Fanuc TP program (LS listing): PgProg.LS

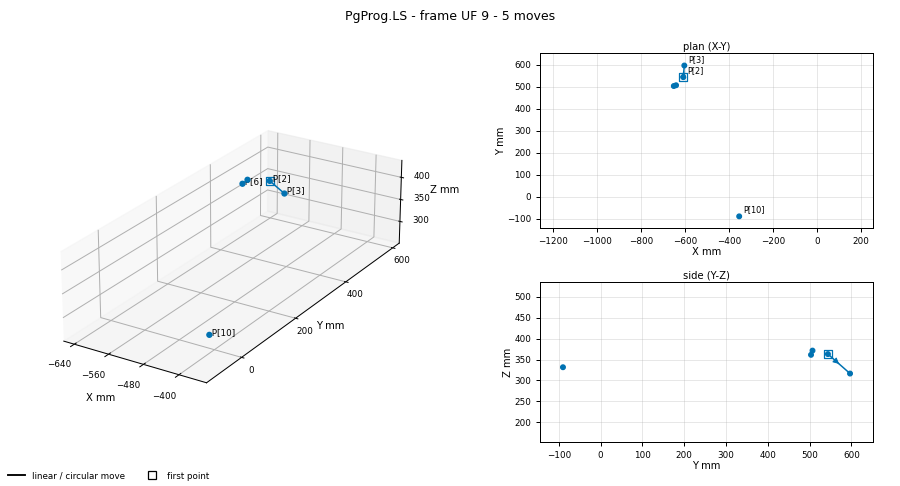
[picture p0: tool path of PgProg.LS in frame UF 9, 5 of 9 moves have a stored position in this frame; points joined in program order, loops and branches not executed]
/PROG  PgProg
/ATTR
OWNER		= MNEDITOR;
COMMENT		= "RoboDK sequence";
PROG_SIZE	= 0;
CREATE		= DATE 31-12-14  TIME 12:00:00;
MODIFIED	= DATE 31-12-14  TIME 12:00:00;
FILE_NAME	= PgProg;
VERSION		= 0;
LINE_COUNT	= 52;
MEMORY_SIZE	= 0;
PROTECT		= READ_WRITE;
TCD:  STACK_SIZE	= 0,
      TASK_PRIORITY	= 50,
      TIME_SLICE	= 0,
      BUSY_LAMP_OFF	= 0,
      ABORT_REQUEST	= 0,
      PAUSE_REQUEST	= 0;
DEFAULT_GROUP	= 1,*,*,*,*;
CONTROL_CODE	= 00000000 00000000;
/MN
   1:  ! Program generated by RoboDK v6.0.7 for Fanuc M-1iA/0.5S on XX ;
   2:  ! /XX/XXXX 18:00:00 ;
   3:  ! Using nominal kinematics. ;
   4:  PR[9,1]=1234.570 ;
   5:  PR[9,2]=-98.765 ;
   6:  PR[9,3]=50.500 ;
   7:  PR[9,4]=0.000 ;
   8:  PR[9,5]=0.000 ;
   9:  PR[9,6]=30.000 ;
  10:  UFRAME[9]=PR[9] ;
  11:  UFRAME_NUM=9 ;
  12:  PR[9,1]=10.000 ;
  13:  PR[9,2]=20.000 ;
  14:  PR[9,3]=150.000 ;
  15:  PR[9,4]=15.000 ;
  16:  PR[9,5]=0.000 ;
  17:  PR[9,6]=0.000 ;
  18:  UTOOL[9]=PR[9] ;
  19:  UTOOL_NUM=9 ;
  20:J P[1] 5% CNT5 ;
  21:L P[2] 250mm/sec CNT5 ;
  22:C P[3]
       P[4] 250mm/sec CNT5 ;
  23:J P[5] 5% CNT5 ;
  24:L P[6] 100mm/sec CNT5 ACC100 ;
  25:L P[7] 100mm/sec CNT0 ACC100 ;
  26:  WAIT  0.50(sec) ;
  27:  PAUSE ;
  28:  MESSAGE[Hello from postgen] ;
  29:  ! a comment ;
  30:  CALL SubProgr ;
  31:  CustomCode(42);
  32:  ThreadProg;
  33:  DO[1]=ON ;
  34:  Valve=OFF ;
  35:  AO[3]=(2.5) ;
  36:  WAIT DI[2]=ON ;
  37:  $WAITTMOUT=1500 ;
  38:  WAIT DI[4]=OFF TIMEOUT, LBL[1] ;
  39:  MESSAGE[Timed out for LBL 1] ;
  40:  PAUSE ;
  41:  LBL[1] ;
  42:  PR[9,1]=0.000 ;
  43:  PR[9,2]=0.000 ;
  44:  PR[9,3]=200.000 ;
  45:  PR[9,4]=0.000 ;
  46:  PR[9,5]=0.000 ;
  47:  PR[9,6]=0.000 ;
  48:  UTOOL[9]=PR[9] ;
  49:  UTOOL_NUM=9 ;
  50:J P[8] 2% CNT0 ACC100 ;
  51:J P[9] 2% CNT0 ACC100 ;
  52:L P[10] 100mm/sec CNT0 ACC100 ;
/POS
P[1]{
   GP1:
    UF : 9, UT : 9,
	J1=    10.000000 deg,	J2=    -20.000000 deg,	J3=    50.000000  mm,
	J4=    30.000000 deg
};
P[2]{
   GP1:
    UF : 9, UT : 9,        CONFIG : 'L, 0, 0, 0',
	X =  -607.850  mm,	Y =   543.849  mm,	Z =   363.215  mm,
	W =  -165.000 deg,	P =    50.000 deg,	R =   150.000 deg
};
P[3]{
   GP1:
    UF : 9, UT : 9,        CONFIG : 'L, 0, 0, 0',
	X =  -602.951  mm,	Y =   596.788  mm,	Z =   316.595  mm,
	W =  -165.000 deg,	P =    50.000 deg,	R =   150.000 deg
};
P[4]{
   GP1:
    UF : 9, UT : 9,        CONFIG : 'L, 0, 0, 0',
	X =  -663.517  mm,	Y =   575.988  mm,	Z =   286.611  mm,
	W =  -165.000 deg,	P =    50.000 deg,	R =   150.000 deg
};
P[5]{
   GP1:
    UF : 9, UT : 9,
	J1=    30.000000 deg,	J2=    25.000000 deg,	J3=    80.000000  mm,
	J4=    -45.000000 deg
};
P[6]{
   GP1:
    UF : 9, UT : 9,        CONFIG : 'L, 0, 0, 0',
	X =  -650.861  mm,	Y =   503.437  mm,	Z =   361.399  mm,
	W =  -165.000 deg,	P =    50.000 deg,	R =   150.000 deg
};
P[7]{
   GP1:
    UF : 9, UT : 9,        CONFIG : 'L, 0, 0, 0',
	X =  -640.584  mm,	Y =   506.980  mm,	Z =   371.534  mm,
	W =  -165.000 deg,	P =    50.000 deg,	R =   150.000 deg
};
P[8]{
   GP1:
    UF : 9, UT : 9,
	J1=    10.000000 deg,	J2=    -20.000000 deg,	J3=    50.000000  mm,
	J4=    30.000000 deg
};
P[9]{
   GP1:
    UF : 9, UT : 9,
	J1=    20.000000 deg,	J2=    -15.000000 deg,	J3=    55.000000  mm,
	J4=    35.000000 deg
};
P[10]{
   GP1:
    UF : 9, UT : 9,        CONFIG : 'L, 0, 0, 0',
	X =  -353.026  mm,	Y =   -90.135  mm,	Z =   331.702  mm,
	W =  -169.444 deg,	P =    40.650 deg,	R =   178.023 deg
};
/END
